Fanuc KAREL source: NC0002.KL

-- PROVISIONAL review KL for V1013-1; original PC SHA256 818b3d47d0b74fb09c1597053c51282c42cfc015785dbabf7e299ffb90e042d4
-- Incomplete behavior may be omitted. Consult companion uncertainty JSON. Do not deploy.
PROGRAM NC0002
%NOLOCKGROUP
-- UNRESOLVED_LOCAL_POOL 1 cells at code offset 3; source declarations unknown
-- DIRECT_LOCAL_WORD_ACCESS alone does not prove INTEGER, REAL, or BOOLEAN
BEGIN
  -- UNRESOLVED_PC offsets 0-8; opcodes 2B,2C,7B
  -- UNRESOLVED_PC offsets 13-20; opcodes 9D,23
  -- UNRESOLVED_PC offsets 25-38; opcodes 21,9D,57,79
  -- UNRESOLVED_PC offsets 43-57; opcodes 21,9D,52,23
  -- UNRESOLVED_PC offsets 62-67; opcodes 7A
  -- UNRESOLVED_PC offsets 72-90; opcodes 21,2E,52,23
  -- UNRESOLVED_PC offsets 100-104; opcodes 7F
  -- UNRESOLVED_PC offsets 109-113; opcodes 27,AA
  -- UNRESOLVED_PC offsets 118-122; opcodes 7F
END NC0002
